FUNCTION F_interpolateTime : REAL
VAR_INPUT
	tX_Old	:	TIME;
	tX_New	:	TIME;
	rY_Old	:	REAL;
	rY_New	:	REAL;
	tX		:	TIME;
END_VAR
VAR
END_VAR

F_interpolateTime	:=	F_interpolateReal(
	rX_Old	:=	F_time2seconds(tX_Old),
	rX_New	:=	F_time2seconds(tX_New),
	rY_Old	:=	rY_Old,
	rY_New	:=	rY_New,
	rX		:=	F_time2seconds(tX)
	);

END_FUNCTION

(* stored: Version 1.1.0.1, ProductVersion 3.1.4024.9
   POU F_interpolateTime: Id {148c1805-e80b-47f2-bb0d-8ebe7a71cd82}, SpecialFunc None *)
